PROGRAM P_COMM_HANDLER
VAR
	i					: UDINT;
	nAddr				: ULINT;
	stReceivedFrom		: ST_UDPFrameEntry;
	sLoggedMessage		: UDP_DATA;
	dVal_1				: LREAL;
	dVal_2				: LREAL;	
	sTurbineData		: S_TURBINEDATA;
	iTemp				: ULINT;
	
	sTxTimer			: TON;
	bSend				: BOOL := FALSE;
	cTxTimerPeriod		: TIME := T#500MS;
	sTurbineCmd			: S_TURBINECMD;
	stSendTo			: ST_UDPFrameEntry;;
END_VAR


(* First we pop from the UDP RX buffer, and process the received data accordingly *)
REPEAT
	fbRxFIFO.RemoveHead( );
	IF fbRxFIFO.bOk THEN

		(* TODO:: Implement received frame handler *)
		stReceivedFrom := fbRxFIFO.stGet;
		IF stReceivedFrom.stRemoteAddr.sAddr = sRemoteHost AND stReceivedFrom.stRemoteAddr.nPort = nRemoteTxPort THEN
// 			sLoggedMessage := stReceivedFrom.sMessage;
			nAddr := 0;
			FOR i := 1 TO c_nNumTurbines DO
				sTurbineData := ParseTurbineData(ADR(stReceivedFrom.sMessage) + nAddr);
				F_InsertTurbineDataIEC61850(nID := i, sTurbineData := sTurbineData);
				nAddr := nAddr + SIZEOF(S_TURBINEDATA);
			END_FOR
		END_IF
// 		MEMCPY(ADR(dVal_1), ADR(sLoggedMessage), SIZEOF(dVal_1));
// 		MEMCPY(ADR(dVal_2), ADR(sLoggedMessage) + SIZEOF(dVal_1), SIZEOF(dVal_2));
// 			ADSLOGSTR( ADSLOG_MSGTYPE_HINT OR ADSLOG_MSGTYPE_LOG OR ADSLOG_MSGTYPE_MSGBOX, '%s', stReceivedFrom.sMessage );
		
	END_IF
UNTIL NOT fbRxFIFO.bOk
END_REPEAT


(* Second, we take the turbine setpoints and transmit to the turbine *)
bSend := sTxTimer.Q;
sTxTimer(IN := NOT sTxTimer.Q, PT := cTxTimerPeriod);

IF bSend THEN
	sTurbineCmd := F_CreateTurbineCMD();
	fbTXFIFO.AddTail( );
	iTemp :=  SIZEOF(sTurbineCmd);
	MEMCPY(ADR(stSendTo.sMessage), ADR(sTurbineCmd), SIZEOF(sTurbineCmd));
	stSendTo.stRemoteAddr.sAddr := sRemoteHost;	(* Remote host IP address *)
	stSendTo.stRemoteAddr.nPort := nRemoteRxPort;	(* Remote host port number *)
	fbTxFIFO.AddTail( stPut := stSendTo );
END_IF

END_PROGRAM

(* stored: Version 1.1.0.1
   POU P_COMM_HANDLER: Id {e2c46c32-4353-43a4-9fe3-574824d63608}, SpecialFunc None *)
